// Tampon circulaire de traces lu par la HMI depuis le dernier nSeq reçu (docs/05 § 9)
FUNCTION_BLOCK FB_TraceBuffer
VAR
    _refBuf : REFERENCE TO ST_TraceBuffer;
END_VAR

METHOD Bind
VAR_INPUT
    refBuf : REFERENCE TO ST_TraceBuffer;
END_VAR
_refBuf REF= refBuf;
END_METHOD

METHOD Add : UDINT
VAR_INPUT
    stTrace : ST_TraceRecord;
END_VAR
VAR
    k : INT;
END_VAR
IF NOT __ISVALIDREF(_refBuf) THEN RETURN; END_IF
_refBuf.nWriteSeq := _refBuf.nWriteSeq + 1;
k := UDINT_TO_INT(_refBuf.nWriteSeq MOD INT_TO_UDINT(GVL_Const.TRACE_BUFFER));
_refBuf.aTrace[k] := stTrace;
_refBuf.aTrace[k].nSeq := _refBuf.nWriteSeq;
Add := _refBuf.nWriteSeq;
END_METHOD

END_FUNCTION_BLOCK

(* stored: Version 1.1.0.1, ProductVersion 3.1.4024.12
   POU FB_TraceBuffer: Id {c16340b6-71d3-5982-9e22-547b6718049b}, SpecialFunc None
   Method Bind: Id {29c60252-8be7-5bb2-afa0-030d01edac96}
   Method Add: Id {a2450718-5112-597e-9d3e-5729c1c866ed} *)
